(* IEC 61131-3 sources: iolistgen/tools/tests/fixtures/sample/src/DUTs, 3 files *)

(* ---- E_DeviceMode.dut.st ---- *)
{attribute 'qualified_only'}
{attribute 'strict'}
// Режим работы устройства (docs/ARCHITECTURE.md, раздел «Режимы»)
TYPE E_DeviceMode :
(
    Auto := 0,          // автоматический
    Manual := 1,        // ручной с HMI
    Local := 2,         // местный пост
    OutOfService := 3   // выведен из работы
) INT;
END_TYPE

(* ---- E_NamurStatus.dut.st ---- *)
{attribute 'qualified_only'}
// Статус диагностики по NAMUR NE 107 (названия — сверить с источником)
TYPE E_NamurStatus :
(
    Good,
    CheckFunction,
    OutOfSpecification,
    MaintenanceRequired,
    Failure
);
END_TYPE

(* ---- U_RawValue.dut.st ---- *)
// Сырое значение из регистра Modbus: как DWORD или как REAL
TYPE U_RawValue :
UNION
    dwRaw : DWORD;
    rValue : REAL;
END_UNION
END_TYPE
